FUNCTION_BLOCK FB_AxisControl
// 单轴基础控制：使能、复位、手动点动、标准回原、停止及反馈。
// 四轴分别使用独立实例；本块不读取位置表，轨迹块通过 xGroupBusy 占用轴控制。
VAR_INPUT
    xPermit : BOOL; // 普通运行及控制权许可；FALSE 请求停车，并禁止新使能和新手动动作。
    xPositiveLimit : BOOL; // 正向硬限位，TRUE 表示触发。
    xNegativeLimit : BOOL; // 负向硬限位，TRUE 表示触发。
    xHomeSensor : BOOL; // 实际原点开关，作为标准回原校准凸轮信号。
    xGroupBusy : BOOL; // 轨迹占用时禁止手动点动、回原和复位抢占。
    Config : ST_AxisConfig; // 本轴行程及动态参数，单位跟随 NC。
END_VAR
VAR_IN_OUT
    Axis : AXIS_REF; // 对应 NC 轴引用，直接操作原轴接口。
    Data : ST_AxisAds; // 内部轴命令及反馈；命令由命令门转交，本块读取命令并更新实际反馈。
END_VAR
VAR
    fbPower : MC_Power; // 轴软件使能实例；Status 才是实际使能反馈，Data.xStart 仅为请求。
    fbJog : MC_Jog; // 正反点动实例；速度单位为 NC 位置单位/秒。
    fbHome : MC_Home; // NC 标准回零实例，使用配置的回零方式和原点凸轮信号。
    fbStop : MC_Stop; // 单轴减速停止实例；Execute 释放后仍需等待 Busy 解锁。
    fbReset : MC_Reset; // NC 轴报警复位实例，不代替运动块或轨迹组的独立故障复位。
    rtHome : R_TRIG; // 回零请求上升沿检测，输入保持 TRUE 不重复发起回零。
    rtReset : R_TRIG; // 轴复位请求上升沿检测，输入保持 TRUE 不重复发起复位。
    xPositionValid : BOOL; // 位置范围单独校验，只用于方向限制。
    xConfigValid : BOOL; // 运动参数校验，只限制点动/回原，不限制基础使能。
    xManual : BOOL; // 允许手动运动的公共条件。
    xStopRequest : BOOL; // 停止、撤使能、许可丢失、限位或运动中参数失效产生的停车条件。
    xHoldPower : BOOL; // 运动/停车未完成或组仍占用时，临时保持已有使能。
    xJogArmed : BOOL; // 联停或轨迹占用后，须先释放按钮才重新允许点动。
    xJogSpeedValid : BOOL; // 点动速度为正且不超过最大速度。
    lrJogVelocity : LREAL; // 本扫描合法点动速度，单位为 NC 位置单位/秒；无效输入置零。
    lrStopDeceleration : LREAL; // 本扫描停车减速度，单位为 NC 位置单位/秒²；参数无效时按 MC_Stop 默认规则处理。
END_VAR

// ReadStatus 在 MAIN 开头统一执行，所有轴使用本周期反馈。
// 1. 回原/复位取上升沿；输入保持 TRUE 不会每扫描重复发起。
rtHome(CLK := Data.gohome);
rtReset(CLK := Data.reset);
// Config 由 MAIN 传入 GVL_motion.aConfig；本块只读取，不覆盖输入参数。
// 2. 分开校验位置和运动参数；未配置时可以基础使能，但不允许发起运动。
xPositionValid := F_AxisPositionValid(Config);
xConfigValid := F_AxisConfigValid(Config);

// 3. 软件使能：Data.xStart 是持续使能请求，xPermit 和有效 I/O 决定能否接受该请求。
// 已经使能的轴在运动、轨迹占用或 MC_Stop 尚未结束时，由 xHoldPower 暂时保持使能。
// MC_Power 先执行，下面的 MC_Stop 使用本扫描更新后的使能反馈。
xHoldPower := fbPower.Status AND (Axis.Status.Moving OR xGroupBusy
    OR (fbStop.Busy AND NOT fbStop.Done AND NOT fbStop.Error));
// 正负方向受硬限位约束，位置范围有效时再检查位置边界。
fbPower(Axis := Axis, Enable := (Data.xStart AND xPermit AND NOT Axis.Status.IoDataInvalid) OR xHoldPower,
    Enable_Positive := NOT xPositiveLimit AND (NOT xPositionValid OR (Axis.NcToPlc.ActPos < Config.lrMaxPosition)),
    Enable_Negative := NOT xNegativeLimit AND (NOT xPositionValid OR (Axis.NcToPlc.ActPos > Config.lrMinPosition)), Override := 100);

// 4. 停车请求：停止、撤使能、许可丢失、限位或运动中参数失效。
xStopRequest := Data.xStop OR NOT Data.xStart OR NOT xPermit OR xPositiveLimit OR xNegativeLimit
    OR (NOT xConfigValid AND (Axis.Status.Moving OR fbJog.Busy OR fbHome.Busy));
// 配置无效也必须能停车；0 按 MC_Stop 默认规则沿用最近运动命令的减速度。
lrStopDeceleration := 0;
IF xConfigValid THEN lrStopDeceleration := Config.lrStopDeceleration; END_IF
// 轨迹占用或外部给定仍开启时，由轨迹块负责停车。
// MC_Stop 的 Execute 释放后，等 Busy 变为 FALSE 才允许新的手动运动。
fbStop(Axis := Axis, Execute := xStopRequest AND fbPower.Status
    AND NOT xGroupBusy AND NOT Axis.Status.ExtSetPointGenEnabled,
    Deceleration := lrStopDeceleration);

// 5. 新手动动作许可：本扫描的使能、停车和反馈状态共同决定能否点动或回原。
// Data.reset 同时阻断手动，避免同一扫描复位和点动并发。
xManual := xPermit AND xConfigValid AND fbPower.Status AND NOT xStopRequest
    AND NOT xGroupBusy AND NOT Axis.Status.ExtSetPointGenEnabled
    AND NOT fbStop.Busy AND NOT Axis.Status.Error AND NOT Axis.Status.IoDataInvalid
    AND NOT fbReset.Busy AND NOT Data.reset;
// 6. 上位机主动复位；本块不自动反复复位故障轴。
fbReset(Axis := Axis, Execute := rtReset.Q AND NOT xGroupBusy
    AND NOT Axis.Status.Moving AND NOT Data.xStop);
// 7. MC_DefaultHoming 使用 NC 配置的回原方式、速度和参考位置。
// 原点输入接实际传感器；点动按钮释放且点动块不忙时才允许启动回原。
fbHome(Axis := Axis, Execute := rtHome.Q AND xManual
    AND NOT fbJog.Busy AND NOT Data.jogz AND NOT Data.jogf,
    HomingMode := MC_DefaultHoming, bCalibrationCam := xHomeSensor);
// 正反同时按下不点动；释放按钮由 MC_Jog 按 NC 参数减速。
// 联停或轨迹占用后，必须先释放点动按钮，防止旧命令自动恢复运动。
IF NOT xManual OR fbHome.Busy THEN xJogArmed := FALSE;
ELSIF NOT Data.jogz AND NOT Data.jogf THEN xJogArmed := TRUE;
END_IF
xJogSpeedValid := (Data.lrJogSpeed > 0) AND (Data.lrJogSpeed <= Config.lrMaxVelocity);
lrJogVelocity := 0;
IF xJogSpeedValid THEN lrJogVelocity := Data.lrJogSpeed; END_IF
// 8. jogz 正向、jogf 负向，保持运行、释放减速；正反同时按下不运行。
// CONTINOUS 是 Tc2_MC2 的实际枚举名称，采用这里传入的速度和动态参数。
fbJog(Axis := Axis, JogForward := Data.jogz AND NOT Data.jogf
    AND xManual AND xJogArmed AND xJogSpeedValid AND NOT fbHome.Busy AND NOT Data.gohome,
    JogBackwards := Data.jogf AND NOT Data.jogz
    AND xManual AND xJogArmed AND xJogSpeedValid AND NOT fbHome.Busy AND NOT Data.gohome,
    Mode := MC_JOGMODE_CONTINOUS, // Tc2_MC2 的枚举名称使用 CONTINOUS 拼写。
    Velocity := lrJogVelocity,
    Acceleration := Config.lrMaxAcceleration, Deceleration := Config.lrStopDeceleration);

// 9. 反馈来源为 NC 实际状态和 MC 输出，不用上位机请求位代替执行结果。
// xEnabled=Power.Status，xHomed=NC.Homed；ErrorID 依 NC/Power/Stop/Home/Jog/Reset 顺序取首项。
Data.lrActualPosition := Axis.NcToPlc.ActPos;
Data.lrSpeed := Axis.NcToPlc.ActVelo;
Data.xMotorRun := Axis.Status.Moving;
Data.xEnabled := fbPower.Status;
Data.xHomed := Axis.Status.Homed;
Data.xPositiveLimit := xPositiveLimit OR Axis.Status.SoftLimitMaxExceeded;
Data.xNegativeLimit := xNegativeLimit OR Axis.Status.SoftLimitMinExceeded;
Data.xOriginSignal := xHomeSensor;
// MC_Stop Execute 保持时 Busy 可持续为 TRUE；停车确认与块释放分开反馈。
Data.xStopped := NOT Axis.Status.Moving AND NOT Axis.Status.IoDataInvalid
    AND (ABS(Axis.NcToPlc.ActVelo) <= 0.000001) AND NOT fbJog.Busy AND NOT fbHome.Busy
    AND NOT fbReset.Busy AND (NOT fbStop.Busy OR fbStop.Done);
Data.xBusy := xGroupBusy OR fbJog.Busy OR fbHome.Busy OR fbStop.Busy OR fbReset.Busy;
Data.udiErrorId := 0;
IF Axis.Status.Error THEN Data.udiErrorId := Axis.Status.ErrorId;
ELSIF fbPower.Error THEN Data.udiErrorId := fbPower.ErrorID;
ELSIF fbStop.Error THEN Data.udiErrorId := fbStop.ErrorID;
ELSIF fbHome.Error THEN Data.udiErrorId := fbHome.ErrorID;
ELSIF fbJog.Error THEN Data.udiErrorId := fbJog.ErrorID;
ELSIF fbReset.Error THEN Data.udiErrorId := fbReset.ErrorID;
END_IF
Data.xError := Axis.Status.Error OR fbPower.Error OR fbStop.Error
    OR fbHome.Error OR fbJog.Error OR fbReset.Error;

END_FUNCTION_BLOCK

(* stored: Version 1.1.0.1
   POU FB_AxisControl: Id {9B2140E4-2674-461A-AEA8-E3B7301EB2D3}, SpecialFunc None *)
